Staubli VAL3: click_refresh.pgx

program click_refresh()
begin
  call initMsg()
  call rs:getLog(sRobotMsg,nMsgType)
end
